// Generated by voz_llm_plc_agent
// Target: Siemens TIA Portal V18 - SCL external source
// Review and compile before any download to physical hardware.

FUNCTION_BLOCK "PLC_PRG"
{ S7_Optimized_Access := 'TRUE' }
VERSION : 0.1
VAR_INPUT
   I_Emergency : Bool := FALSE;
   I_Automatic_Motor_Command : Bool := FALSE;
   I_Mode_Manual : Bool := FALSE;
   I_Manual_Motor_Command : Bool := FALSE;
END_VAR
VAR_OUTPUT
   Q_Motor_Enable : Bool := FALSE;
END_VAR
VAR
   M_AutoMode : Bool;
   M_ManualMode : Bool;
END_VAR
BEGIN
(* Seleccion de modo de operacion (excluyentes) *)
#M_AutoMode := #I_Mode_Manual;
#M_ManualMode := NOT #I_Mode_Manual;
(* Salidas: contribucion automatica (secuencia/condiciones) y manual, con sus bloqueos *)
#Q_Motor_Enable := ((#M_AutoMode AND #I_Automatic_Motor_Command AND NOT #I_Emergency) OR (#M_ManualMode AND #I_Manual_Motor_Command AND (#M_ManualMode))) AND NOT #I_Emergency;
(* Bloqueo: #I_Emergency fuerza a FALSE #Q_Motor_Enable de inmediato *)
IF #I_Emergency THEN
    #Q_Motor_Enable := FALSE;
END_IF;
END_FUNCTION_BLOCK

DATA_BLOCK "DB_PLC_PRG"
{ S7_Optimized_Access := 'TRUE' }
VERSION : 0.1
NON_RETAIN
"PLC_PRG"
BEGIN
END_DATA_BLOCK

ORGANIZATION_BLOCK "Main"
{ S7_Optimized_Access := 'TRUE' }
VERSION : 0.1
BEGIN
   "DB_PLC_PRG"(
      I_Emergency := "I_Emergency",
      I_Automatic_Motor_Command := "I_Automatic_Motor_Command",
      Q_Motor_Enable => "Q_Motor_Enable",
      I_Mode_Manual := "I_Mode_Manual",
      I_Manual_Motor_Command := "I_Manual_Motor_Command"
   );
END_ORGANIZATION_BLOCK
